// TIA Portal V21 export
// export: Created 2026-11-11T00:47:54.6425213Z, ExportSetting WithDefaults, DisplayName Totally Integrated Automation Portal, DisplayVersion V21 Update 3, DisplayName STEP 7 Professional, DisplayVersion V21 Update 3, DisplayName STEP 7 Safety, DisplayVersion V21, DisplayName Tech WebApplication, DisplayVersion V21, DisplayName WinCC Basic/Comfort/Advanced, DisplayVersion V21 Update 3, DisplayName WinCC Unified, DisplayVersion V21 Update 3
FUNCTION_BLOCK "FB_Lad_ex159"   // FB210, LAD
{ S7_Optimized_Access := 'TRUE' }
VERSION : 0.1
// stored: AutoNumber true, IsIECCheckEnabled false, IsRetainMemResEnabled false, MemoryReserve 100, SetENOAutomatically false, UDAEnableTagReadback false
   VAR_INPUT
      v_ioid : Byte;
      v_laddr : HW_ANY;
   END_VAR
   VAR_OUTPUT
      v_ret_val : Int;
      v_pecount : Int;
      v_pacount : Int;
   END_VAR
BEGIN

REGION Network 1: RD_LGADR - Determine IO addresses from the hardware identifier
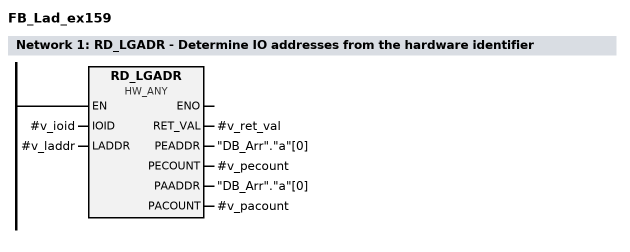
   RUNG wire#powerrail
      { S7_Templates := "laddr_type := HW_ANY" } RD_LGADR(IOID := #v_ioid, LADDR := #v_laddr, RET_VAL => #v_ret_val, PEADDR => "DB_Arr"."a"[0], PECOUNT => #v_pecount, PAADDR => "DB_Arr"."a"[0], PACOUNT => #v_pacount)
   END_RUNG
   // the same network as SCL:
   #v_ret_val := RD_LGADR(IOID := #v_ioid,
                          LADDR := #v_laddr,
                          PEADDR => "DB_Arr"."a"[0],
                          PECOUNT => #v_pecount,
                          PAADDR => "DB_Arr"."a"[0],
                          PACOUNT => #v_pacount);
END_REGION
END_FUNCTION_BLOCK
